Fanuc KAREL source: kt00010.KL

PROGRAM KT00010
%NOLOCKGROUP
VAR
R1:REAL;I2:INTEGER;OUT:REAL
BEGIN
--
--
R1=2.0
I2=3
OUT=(R1+(I2))
END KT00010
